(*
SPDX-FileCopyrightText: © 2026 Oleksandr Tiutyk <trofimich@gmail.com>
SPDX-License-Identifier: MIT
License: https://opensource.org/license/mit
*)
(*!
<summary>Selects the deliberate backend outcome used by logger containment tests.</summary>
*)
{attribute 'qualified_only'}
{attribute 'strict'}
TYPE LOGGER_DELIVERY_BEHAVIOR :
(
	ACCEPT,
	REFUSE,
	THROW_EXCEPTION
);
END_TYPE

(* stored: Version 1.1.0.1
   DUT LOGGER_DELIVERY_BEHAVIOR: Id {c9a41943-8193-4e71-8db8-c189581f7f7c} *)
